SUBAPPLICATION Uebung_147 (* Übung zu DlPgnSend: PropA einmal mit 20 Byte global senden, ohne install *)
  (* Standard: 61499-2; Description: Copyright (c) 2026 Meisterschulen am Ostbahnhof This program and the accompanying materials are made available under the terms of the Eclipse Public License 2.0 which is available at https://www.eclipse.org/legal/epl-2.0/ SPDX-License-Identifier: EPL-2.0 *)
  (* Version 1.0, 2026-11-17, Franz Höpfinger, Meisterschulen am Ostbahnhof, initial API and implementation and/or initial documentation *)
  PACKAGE Uebungen;
  IMPORT Uebungen::const::Uebung_120_129::Filter::ADD_ALL_PASS;
  IMPORT Uebungen::const::Uebung_120_129::Filter::FLT_ALL_PASS;
  IMPORT isobus::pgn::ISOUSERHOME_e::thisMember;
  IMPORT isobus::pgn::ISO_CAN_NODE::NODE1;
  IMPORT isobus::pgn::const::PgnDef::PGN_PDU1_PropA;
  IMPORT logiBUS::io::DI::logiBUS_DI::Input_I1;
  IMPORT logiBUS::io::DI::logiBUS_DI_Events::BUTTON_SINGLE_CLICK;
  IMPORT isobus::pgn::HANDLE::GLOBAL;
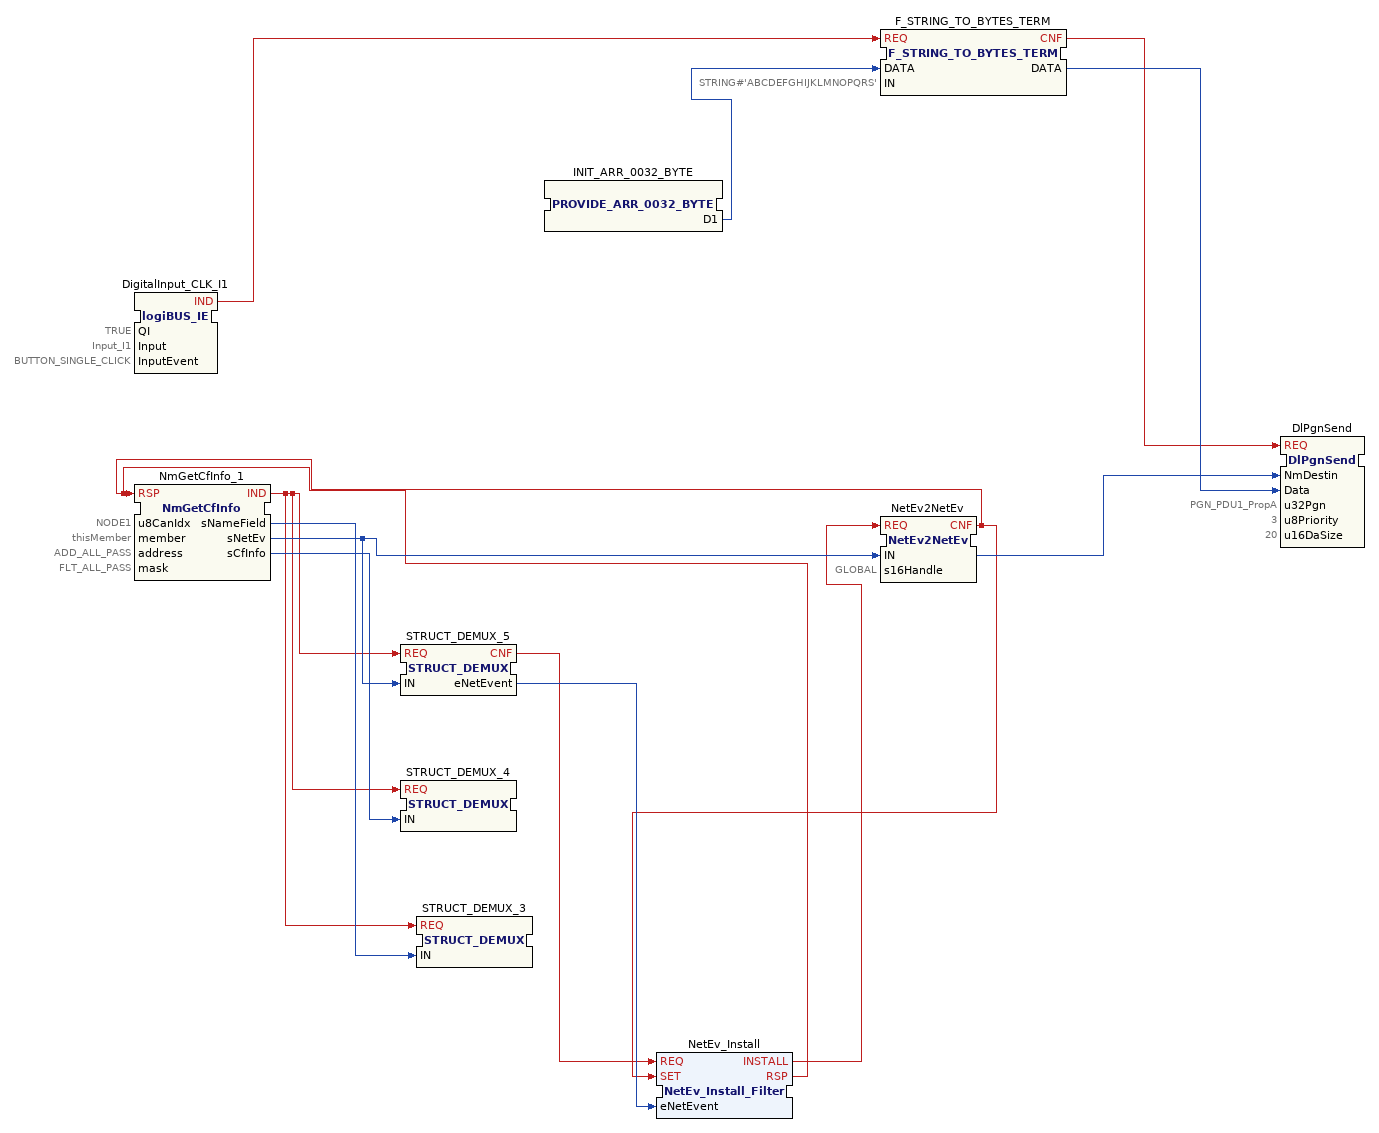
  (* DlPgnSend: eine PGN einmal senden, ohne install NmDestin aus der eigenen CF (thisMember, Active): s16OwnCfHnd = Sender, s16Handle = HANDLE::GLOBAL. I1 Klick: PropA (0xEF00) mit 20 Byte (A-S + 16#00) global, mehr als 8 Byte = TP BAM. s16Status 0 = OK. Empfänger: Übung 139 zeigt den Text. *)
  FBS
    STRUCT_DEMUX_3 : eclipse4diac::convert::STRUCT_DEMUX; {SET_ATTRIBUTE(StructuredType, isobus::pgn::NAMEFIELD_T)}
    NmGetCfInfo_1 : isobus::pgn::NmGetCfInfo(u8CanIdx := NODE1, member := thisMember, address := ADD_ALL_PASS, mask := FLT_ALL_PASS);
    STRUCT_DEMUX_4 : eclipse4diac::convert::STRUCT_DEMUX; {SET_ATTRIBUTE(StructuredType, isobus::pgn::CF_INFO_T)}
    STRUCT_DEMUX_5 : eclipse4diac::convert::STRUCT_DEMUX; {SET_ATTRIBUTE(StructuredType, isobus::pgn::ISONETEVENT_T)}
    NetEv2NetEv : isobus::pgn::NetEv2NetEv(s16Handle := GLOBAL);
    INIT_ARR_0032_BYTE : eclipse4diac::convert::providers::PROVIDE_ARR_0032_BYTE;
    F_STRING_TO_BYTES_TERM : logiBUS::utils::dyn_arr::F_STRING_TO_BYTES_TERM(IN := STRING#'ABCDEFGHIJKLMNOPQRS');
    DigitalInput_CLK_I1 : logiBUS::io::DI::logiBUS_IE(QI := TRUE, Input := Input_I1, InputEvent := BUTTON_SINGLE_CLICK);
    DlPgnSend : isobus::pgn::tx::DlPgnSend(u32Pgn := PGN_PDU1_PropA, u8Priority := 3, u16DaSize := 20); (* einmal senden, ohne install *)
  END_FBS
  SUBAPPS
    NetEv_Install : MyLib::sys::NetEv_Install_Filter;
  END_SUBAPPS
  EVENT_CONNECTIONS
    NmGetCfInfo_1.IND TO STRUCT_DEMUX_3.REQ;
    NmGetCfInfo_1.IND TO STRUCT_DEMUX_4.REQ;
    NmGetCfInfo_1.IND TO STRUCT_DEMUX_5.REQ;
    DigitalInput_CLK_I1.IND TO F_STRING_TO_BYTES_TERM.REQ;
    STRUCT_DEMUX_5.CNF TO NetEv_Install.REQ;
    NetEv_Install.INSTALL TO NetEv2NetEv.REQ;
    NetEv_Install.RSP TO NmGetCfInfo_1.RSP;
    NetEv2NetEv.CNF TO NetEv_Install.SET;
    NetEv2NetEv.CNF TO NmGetCfInfo_1.RSP;
    F_STRING_TO_BYTES_TERM.CNF TO DlPgnSend.REQ;
  END_CONNECTIONS
  DATA_CONNECTIONS
    NmGetCfInfo_1.sNameField TO STRUCT_DEMUX_3.IN;
    NmGetCfInfo_1.sNetEv TO STRUCT_DEMUX_5.IN;
    NmGetCfInfo_1.sCfInfo TO STRUCT_DEMUX_4.IN;
    NmGetCfInfo_1.sNetEv TO NetEv2NetEv.IN;
    INIT_ARR_0032_BYTE.D1 TO F_STRING_TO_BYTES_TERM.DATA;
    STRUCT_DEMUX_5.eNetEvent TO NetEv_Install.eNetEvent;
    NetEv2NetEv. TO DlPgnSend.NmDestin;
    F_STRING_TO_BYTES_TERM.DATA TO DlPgnSend.Data;
  END_CONNECTIONS
END_SUBAPPLICATION
